(* IEC 61131-3 sources: autonomer-verladearm/plc/codesys, 13 files *)

(* ---- DUT_Pd.st ---- *)
(* Prozessdaten eines MOVITRAC advanced mit MOVIKIT Positioning Drive (Applikationslevel 1, 8 PD).
   Belegung nach Handbuch 33350930 (11/2025), Kap. 8 – im E/A-Abbild des PROFINET-Geräts auf
   diese Felder legen. *)
TYPE ST_PdAxis :
STRUCT
    aPA : ARRAY[1..8] OF WORD;   (* SPS -> Umrichter *)
        (* PA1 Steuerwort, PA2 Geschwindigkeit, PA3 Beschleunigung, PA4 Verzögerung,
           PA5 Ausgänge, PA6 Betriebsart (400 = absolut), PA7/PA8 Zielposition (32 Bit, High/Low) *)
    aPE : ARRAY[1..8] OF WORD;   (* Umrichter -> SPS *)
        (* PE1 Statuswort, PE2 Geschwindigkeit, PE3 Fehlercode, PE4 Moment, PE5 Eingänge,
           PE6 aktive Betriebsart, PE7/PE8 Istposition (32 Bit, High/Low) *)
END_STRUCT
END_TYPE

(* ---- GVL_Achsen.st ---- *)
(* Achsen J1..J3: Prozessdaten (im E/A-Abbild der drei MOVITRAC zuordnen), Fahrbefehle und
   Istwerte. Fahrbefehle schreibt immer nur ein Besitzer (Automatik oder Hand). *)
{attribute 'qualified_only'}
VAR_GLOBAL
    aPd        : ARRAY[1..3] OF ST_PdAxis;   (* E/A-Abbild MOVITRAC J1, J2, J3 *)
    (* Befehle *)
    aCmdZiel   : ARRAY[1..3] OF REAL;        (* ° *)
    aCmdV      : ARRAY[1..3] OF REAL;        (* °/s *)
    aCmdA      : ARRAY[1..3] OF REAL;        (* °/s² *)
    xCmdStart  : BOOL;                       (* Flanke = neues Ziel, halten während der Fahrt *)
    xCmdStop   : BOOL;
    xCmdReset  : BOOL;
    iBesitzer  : INT;                        (* 0 frei, 1 Automatik, 2 Hand *)
    (* Istwerte *)
    aIst       : ARRAY[1..3] OF REAL;        (* ° *)
    xAlleBereit: BOOL;
    xAlleInPos : BOOL;
    xAchsFehler: BOOL;
END_VAR

(* ---- GVL_IO.st ---- *)
(* Ein- und Ausgänge. Im Gerätebaum (TwinCAT: E/A-Abbild der EtherCAT-Klemmen bzw. PROFINET-
   Geräte) diesen Variablen zuordnen. Sicherheitssignale kommen als MELDUNG der Sicherheits-
   steuerung (TwinSAFE) – sie schaltet STO selbst, die SPS kann sie nicht überstimmen.
   Not-Halt am Arm schaltet die Pumpe festverdrahtet über die Sicherheitssteuerung ab (nicht hier). *)
{attribute 'qualified_only'}
VAR_GLOBAL
    (* Bedienung am Schaltschrank *)
    xStartTaster      : BOOL;   (* Leuchttaster "Beladen starten" *)
    xQuittTaster      : BOOL;   (* Quittieren *)
    xBetriebsartHand  : BOOL;   (* Schlüsselschalter: TRUE = Hand, FALSE = Automatik *)
    xLampeStart       : BOOL;   (* Lampe im Starttaster *)
    xMeldeGruen       : BOOL;   (* Park / bereit, Fahrzeug darf fahren *)
    xMeldeGelb        : BOOL;   (* Automatik läuft *)
    xMeldeRot         : BOOL;   (* Störung *)

    (* Handbediengerät (Zustimmung wertet die Sicherheitssteuerung aus) *)
    xHandAchse1       : BOOL;
    xHandAchse2       : BOOL;
    xHandAchse3       : BOOL;
    xHandPlus         : BOOL;
    xHandMinus        : BOOL;
    xHandBremseLueften: BOOL;   (* nur J1/J2, Freigabe zusätzlich durch Sicherheitssteuerung *)

    (* Meldungen der Sicherheitssteuerung *)
    xSicherheitOk     : BOOL;   (* kein Not-Halt, STO aufgehoben *)
    xZustimmung       : BOOL;   (* Zustimmtaster Mittelstellung (nur Hand) *)
    xKlapptreppeRuhe  : BOOL;   (* Klapptreppe in Ruhelage *)
    xLichtschranke    : BOOL;   (* Stellplatz belegt *)

    (* Prozess am Arm *)
    xGrenzNass        : BOOL;   (* Grenzschalter Nachziehen, ca. 10–15 cm über Auslassende: nass *)
    xUeberfuellAus    : BOOL;   (* Überfüllsicherung ausgelöst (schaltet die Pumpe selbst ab) *)
    xKlappeAuf        : BOOL;   (* Absperrklappe Rückmeldung auf *)
    xKlappeZu         : BOOL;   (* Absperrklappe Rückmeldung zu *)
    xKlappeOeffnen    : BOOL;   (* Ausgang Absperrklappe (gehört zum Arm) *)

    (* Abtropfsicherung: rein mechanisch, keine Signale (Entscheidung 04.11.2026) *)

    (* Leitstelle (PLS) – Menge, Pumpe und Füllende steuert die Leitstelle; Signale mit BASF
       abstimmen (Mail an BASF 09.11.2026) *)
    xPlsFreigabe      : BOOL;   (* Verladung freigegeben (Auftrag liegt vor) *)
    iPlsProdukt       : INT;
    aPlsDome          : ARRAY[1..4] OF INT;    (* Füllschritte: DomeNo, 0 = automatisch *)
    iPlsSchritte      : INT;    (* Anzahl Füllschritte (Kammern), 1 = Kammern verbunden *)
    xPlsPumpeLaeuft   : BOOL;   (* Rückmeldung: Pumpe läuft *)
    xPlsBefuellEnde   : BOOL;   (* "Befüllung Ende" für den aktuellen Füllschritt (Pumpe aus) *)
    xArmBereit        : BOOL;   (* an PLS: Arm im Tank, Klappe offen – Befüllung freigegeben *)
    xBefuellStoppen   : BOOL;   (* an PLS: Pumpe abschalten (Störung, Maximalhöhe, Arm am Ende) *)
END_VAR

(* ---- GVL_Param.st ---- *)
(* Parameter Prototyp HETA. Werte aus vision/config/anlagen/heta_prototyp.yaml (drives, arm.joints)
   und docs/fuellstand_ueberfuellsicherung.md. Bei der Inbetriebnahme prüfen. *)
{attribute 'qualified_only'}
VAR_GLOBAL CONSTANT
    INTERFACE_VERSION : INT := 3;
    MAX_WP            : INT := 16;
    TIMEOUT_JOB       : TIME := T#5S;       (* Done muss innerhalb 5 s kommen *)
    TIMEOUT_HEARTBEAT : TIME := T#1S;
    TIMEOUT_MOVE_ADD  : TIME := T#10S;      (* Reserve zur berechneten Fahrzeit *)
    BERUHIGEN         : TIME := T#3S;       (* Auslass pendelt frei aus (J4) *)
    ABTROPFEN         : TIME := T#60S;      (* BASF: 1 min reicht oft nicht – mit Abtropfsicherung *)
    FAKTOR_LANGSAM    : REAL := 0.3;        (* Eintauchen, Herausfahren, Nachziehen *)
    FAKTOR_HAND       : REAL := 0.2;        (* Tippen *)
    TOL_POS           : REAL := 0.2;        (* ° Position erreicht *)
    TOL_PARK          : REAL := 0.5;        (* ° in Parkstellung *)
    MAX_KORREKTUR     : REAL := 50.0;       (* mm Job 2, darüber Abbruch *)
    ANFAHRHOEHE       : REAL := 0.3;        (* m über Domrand (arm.approach_height) *)
    (* Nachziehen mit einem Grenzschalter (Stand 09.11.2026) *)
    SENSOR_HOEHE      : REAL := 0.12;       (* m Grenzschalter über Auslassende (10–15 cm) *)
    NACHZIEH_SCHRITT  : REAL := 0.05;       (* m Hub je Schaltvorgang -> Auslass 7–12 cm unter Spiegel *)
    TROCKEN_ZEIT      : TIME := T#10S;      (* nach dem Hub muss der Grenzschalter trocken sein *)
    MAX_OHNE_SCHALTEN : TIME := T#30M;      (* Pumpe läuft, Grenzschalter schaltet nie: Störung *)
    PUMPE_AUSLAUF     : TIME := T#3S;       (* nach "Pumpe aus" warten, dann Klappe zu *)
    PUMPE_AUS_MAX     : TIME := T#15S;      (* Pumpe meldet nicht aus: Klappe trotzdem zu, Störung *)
END_VAR
VAR_GLOBAL
    (* je Achse J1..J3: Höchstgeschwindigkeit [°/s], Beschleunigung [°/s²], Grenzen und Park [°] *)
    aVmax   : ARRAY[1..3] OF REAL := [6.0, 6.0, 5.93];
    aAmax   : ARRAY[1..3] OF REAL := [1.5, 3.0, 3.95];   (* = vmax / Rampe 4 / 2 / 1,5 s *)
    rRuckzeit : REAL := 0.3;                             (* s, auf allen Achsen gleich *)
    aMin    : ARRAY[1..3] OF REAL := [-120.0, -140.0, -45.0];
    aMax    : ARRAY[1..3] OF REAL := [120.0, 140.0, 45.0];
    aPark   : ARRAY[1..3] OF REAL := [70.0, -135.0, 10.0]; (* heta_prototyp.yaml, bei IBN anpassen *)
    (* Eintauchtiefe je Produkt [m unter Domrand], Index = ProductId 0..9 *)
    (* ca. 20 cm über dem Tankboden: Domrand bis Boden 2,10–2,30 m (BASF 24.11.) – flachster Tank 2,10 m *)
    aEintauchtiefe : ARRAY[0..9] OF REAL := [1.9, 1.9, 1.9, 1.9, 1.9, 1.9, 1.9, 1.9, 1.9, 1.9];
    rMaxHoeheUnterRand : REAL := 0.28;   (* m: Füllende Ebene 2, knapp unter der Überfüllsicherung (ca. 0,2 m) *)
END_VAR

(* ---- GVL_Vision.st ---- *)
(* Schnittstelle Vision-PC <-> SPS, InterfaceVersion 3 (docs/schnittstelle.md).
   Gleiche Namen und Datentypen wie DB_Vision (plc/DB_Vision.db), damit der Vision-Dienst ohne
   Codeänderung verbindet. In der Symbolkonfiguration für OPC UA freigeben (Lesen/Schreiben). *)
{attribute 'qualified_only'}
VAR_GLOBAL
    (* SPS -> PC *)
    HeartbeatPLC   : INT;
    Trigger        : BOOL;
    Job            : INT;      (* 1 messen+planen, 2 nachmessen, 3 Rückfahrt, 0 nur messen *)
    ProductId      : INT;
    DomeNo         : INT;      (* 0 automatisch, n = n-ter offener Dom von vorn *)
    Reset          : BOOL;
    ActualJ1       : REAL;     (* Servo-Istwinkel [°] *)
    ActualJ2       : REAL;
    ActualJ3       : REAL;
    AxesHomed      : BOOL;
    ArmState       : INT;      (* 0 Park, 1 fährt, 2 über Dom, 3 eingetaucht, 9 Störung *)
    (* PC -> SPS *)
    HeartbeatPC    : INT;
    Ready          : BOOL;
    Busy           : BOOL;
    Done           : BOOL;
    Error          : BOOL;
    ErrorCode      : INT;
    ResultId       : DINT;
    TargetX        : REAL;     (* mm, Armbasis *)
    TargetY        : REAL;
    TargetZ        : REAL;
    NormalX        : REAL;
    NormalY        : REAL;
    NormalZ        : REAL;
    DiameterMm     : REAL;
    Confidence     : REAL;
    DomeCount      : INT;
    DomeSelected   : INT;
    WaypointCount  : INT;
    WaypointsJ1    : ARRAY[1..16] OF REAL;   (* Servo-Sollwinkel [°] *)
    WaypointsJ2    : ARRAY[1..16] OF REAL;
    WaypointsJ3    : ARRAY[1..16] OF REAL;
    ApproachIndex  : INT;      (* Stützpunkt "über dem Dom", 0 = keiner *)
    CorrectionX    : REAL;     (* mm, Job 2 *)
    CorrectionY    : REAL;
    InterfaceVersion : INT;
END_VAR

(* ---- F_Hilfen.st ---- *)
(* Hilfsfunktionen für den Ablauf. In CODESYS je Funktion ein eigenes Objekt (POU) anlegen. *)

(* ---------------------------------------------------------------------------------------- *)
(* Arm in Parkstellung? *)
FUNCTION F_InPark : BOOL
VAR
    i : INT;
END_VAR
F_InPark := TRUE;
FOR i := 1 TO 3 DO
    IF ABS(GVL_Achsen.aIst[i] - GVL_Param.aPark[i]) > GVL_Param.TOL_PARK THEN
        F_InPark := FALSE;
    END_IF
END_FOR
END_FUNCTION

(* ---------------------------------------------------------------------------------------- *)
(* Höhe des Auslassendes relativ zum Domrand [m] für eine Lage in der Nachzieh-Tabelle.
   Tabelle = Eintauch-Stützpunkte aus Job 2, gleichmäßig von ANFAHRHOEHE über dem Rand (Lage 1)
   bis rTiefe unter dem Rand (Lage iTab). *)
FUNCTION F_Hoehe : REAL
VAR_INPUT
    rPos   : REAL;   (* 1 .. iTab *)
    iTab   : INT;
    rTiefe : REAL;
END_VAR
IF iTab < 2 THEN
    F_Hoehe := GVL_Param.ANFAHRHOEHE;
ELSE
    F_Hoehe := GVL_Param.ANFAHRHOEHE
               - (rPos - 1.0) / INT_TO_REAL(iTab - 1) * (GVL_Param.ANFAHRHOEHE + rTiefe);
END_IF
END_FUNCTION

(* ---------------------------------------------------------------------------------------- *)
(* Umkehrung: Lage in der Tabelle für eine Höhe relativ zum Domrand. *)
FUNCTION F_PosFuerHoehe : REAL
VAR_INPUT
    rHoehe : REAL;
    iTab   : INT;
    rTiefe : REAL;
END_VAR
IF iTab < 2 THEN
    F_PosFuerHoehe := 1.0;
ELSE
    F_PosFuerHoehe := LIMIT(1.0,
        1.0 + (GVL_Param.ANFAHRHOEHE - rHoehe) / (GVL_Param.ANFAHRHOEHE + rTiefe) * INT_TO_REAL(iTab - 1),
        INT_TO_REAL(iTab));
END_IF
END_FUNCTION

(* ---------------------------------------------------------------------------------------- *)
(* Servowinkel einer Achse für eine Lage in der Tabelle: zwischen den Stützpunkten linear im
   Gelenkraum (wie tools/plc_simulator.py table_at). *)
FUNCTION F_TabWinkel : REAL
VAR_INPUT
    rPos   : REAL;
    iTab   : INT;
    iAchse : INT;
END_VAR
VAR_IN_OUT
    aTab   : ARRAY[1..16, 1..3] OF REAL;
END_VAR
VAR
    k : INT;
    u : REAL;
END_VAR
k := LIMIT(1, DINT_TO_INT(TRUNC(rPos)), MAX(iTab - 1, 1));
u := LIMIT(0.0, rPos - INT_TO_REAL(k), 1.0);
IF iTab < 2 THEN
    F_TabWinkel := aTab[1, iAchse];
ELSE
    F_TabWinkel := aTab[k, iAchse] + u * (aTab[k + 1, iAchse] - aTab[k, iAchse]);
END_IF
END_FUNCTION

(* ---- FB_PdAxis.st ---- *)
(* Eine Achse über MOVIKIT Positioning Drive: Ziel, Geschwindigkeit, Beschleunigung vorgeben,
   Istposition und Status lesen. Positionieren, Rampen und Ruckbegrenzung macht der Umrichter.

   !!! Bitbelegung von Steuer- und Statuswort und die Anwendereinheiten vor der Inbetriebnahme
   mit dem SEW-Handbuch (Kap. 8) und MOVISUITE abgleichen – hier als Konstanten mit
   Platzhalterwerten. Anwendereinheit: 1 Inkrement = 0,001° am Gelenk (in MOVISUITE einstellen). *)
FUNCTION_BLOCK FB_PdAxis
VAR_INPUT
    xEnable  : BOOL;          (* Freigabe (STO aufgehoben, keine Störung) *)
    xStart   : BOOL;          (* steigende Flanke: neues Ziel übernehmen *)
    xStop    : BOOL;          (* Halt mit Verzögerung *)
    xReset   : BOOL;          (* Fehler quittieren *)
    rZiel    : REAL;          (* ° *)
    rV       : REAL;          (* °/s *)
    rA       : REAL;          (* °/s² (Beschleunigung = Verzögerung) *)
END_VAR
VAR_OUTPUT
    rIst     : REAL;          (* ° *)
    xBereit  : BOOL;          (* Umrichter bereit / freigegeben *)
    xInPos   : BOOL;          (* Position erreicht *)
    xFehler  : BOOL;
    wFehler  : WORD;
END_VAR
VAR_IN_OUT
    stPd     : ST_PdAxis;
END_VAR
VAR CONSTANT
    EINHEIT_POS    : REAL := 1000.0;     (* Inkremente je ° (Anwendereinheit 0,001°) *)
    EINHEIT_V      : REAL := 100.0;      (* PA2: 0,01 °/s – prüfen *)
    EINHEIT_A      : REAL := 100.0;      (* PA3/PA4: 0,01 °/s² – prüfen *)
    BETRIEBSART_ABS: WORD := 400;
    (* Steuerwort PA1 – PLATZHALTER, laut Handbuch prüfen *)
    CW_FREIGABE    : WORD := 16#0001;
    CW_START       : WORD := 16#0002;
    CW_HALT        : WORD := 16#0004;
    CW_RESET       : WORD := 16#0100;
    (* Statuswort PE1 – PLATZHALTER, laut Handbuch prüfen *)
    SW_BEREIT      : WORD := 16#0001;
    SW_INPOS       : WORD := 16#0004;
    SW_FEHLER      : WORD := 16#0020;
END_VAR
VAR
    rtStart  : R_TRIG;
    dIst     : DINT;
    dZiel    : DINT;
    wStw     : WORD;
END_VAR

rtStart(CLK := xStart);

(* Istwerte *)
dIst := INT_TO_DINT(WORD_TO_INT(stPd.aPE[7])) * 65536 + WORD_TO_DINT(stPd.aPE[8]);   (* High-Wort mit Vorzeichen *)
rIst := DINT_TO_REAL(dIst) / EINHEIT_POS;
xBereit := (stPd.aPE[1] AND SW_BEREIT) <> 0;
xFehler := (stPd.aPE[1] AND SW_FEHLER) <> 0;
wFehler := stPd.aPE[3];

(* Sollwerte: bei neuem Ziel übernehmen *)
IF rtStart.Q THEN
    dZiel := REAL_TO_DINT(rZiel * EINHEIT_POS);
    stPd.aPA[2] := DINT_TO_WORD(LIMIT(1, REAL_TO_DINT(ABS(rV) * EINHEIT_V), 32767));
    stPd.aPA[3] := DINT_TO_WORD(LIMIT(1, REAL_TO_DINT(ABS(rA) * EINHEIT_A), 32767));
    stPd.aPA[4] := stPd.aPA[3];
    stPd.aPA[7] := DWORD_TO_WORD(SHR(DINT_TO_DWORD(dZiel), 16));
    stPd.aPA[8] := DWORD_TO_WORD(DINT_TO_DWORD(dZiel));
END_IF
stPd.aPA[6] := BETRIEBSART_ABS;

wStw := 0;
IF xEnable THEN wStw := wStw OR CW_FREIGABE; END_IF
IF xEnable AND xStart AND NOT xStop THEN wStw := wStw OR CW_START; END_IF
IF xStop THEN wStw := wStw OR CW_HALT; END_IF
IF xReset THEN wStw := wStw OR CW_RESET; END_IF
stPd.aPA[1] := wStw;

xInPos := ((stPd.aPE[1] AND SW_INPOS) <> 0) AND ABS(rIst - rZiel) <= GVL_Param.TOL_POS;

(* ---- FB_SyncMove.st ---- *)
(* Synchrone Fahrt aller drei Achsen zu einem Stützpunkt (docs/schnittstelle.md):
   Die langsamste Achse bestimmt die Fahrzeit; jede Achse bekommt Geschwindigkeit und
   Beschleunigung proportional zu ihrem Weg, gleiche Ruckzeit auf allen Achsen -> alle starten
   und kommen gleichzeitig an, der Arm fährt die geprüfte Gerade im Gelenkraum.
   Gleiche Rechnung wie Drives.sync() in vision/src/verladearm_vision/drives.py. *)
FUNCTION_BLOCK FB_SyncMove
VAR_INPUT
    xExecute : BOOL;                   (* steigende Flanke startet *)
    aZiel    : ARRAY[1..3] OF REAL;    (* ° *)
    rFaktor  : REAL := 1.0;            (* Geschwindigkeitsfaktor, z. B. 0,3 beim Eintauchen *)
    xAbbruch : BOOL;                   (* Halt mit Verzögerung *)
END_VAR
VAR_OUTPUT
    xBusy    : BOOL;
    xDone    : BOOL;
    xError   : BOOL;
    sFehler  : STRING(80);
    rDauer   : REAL;                   (* s, berechnete Fahrzeit *)
END_VAR
VAR
    rtExec   : R_TRIG;
    iSchritt : INT;
    tonZeit  : TON;
    i        : INT;
    d        : ARRAY[1..3] OF REAL;
    rCruise, rPush, rRamp : REAL;
    rFak     : REAL;
END_VAR

rtExec(CLK := xExecute);
IF rtExec.Q THEN
    xDone := FALSE; xError := FALSE; sFehler := '';
    rFak := LIMIT(0.01, rFaktor, 1.0);
    rCruise := 0.0; rPush := 0.0;
    FOR i := 1 TO 3 DO
        aZiel[i] := LIMIT(GVL_Param.aMin[i], aZiel[i], GVL_Param.aMax[i]);   (* Software-Endlagen *)
        d[i] := ABS(aZiel[i] - GVL_Achsen.aIst[i]);
        rCruise := MAX(rCruise, d[i] / (GVL_Param.aVmax[i] * rFak));
        rPush := MAX(rPush, d[i] / GVL_Param.aAmax[i]);
    END_FOR
    IF rPush < 1.0E-6 THEN
        xDone := TRUE; iSchritt := 0;       (* schon am Ziel *)
    ELSE
        IF SQRT(rPush) >= rCruise THEN      (* Dreieck: Höchstgeschwindigkeit nicht erreicht *)
            rCruise := SQRT(rPush); rRamp := rCruise;
        ELSE
            rRamp := rPush / rCruise;
        END_IF
        rDauer := rCruise + rRamp + GVL_Param.rRuckzeit;
        FOR i := 1 TO 3 DO
            GVL_Achsen.aCmdZiel[i] := aZiel[i];
            GVL_Achsen.aCmdV[i] := MAX(d[i] / rCruise, 0.001);
            GVL_Achsen.aCmdA[i] := MAX(d[i] / rCruise / rRamp, 0.001);
        END_FOR
        GVL_Achsen.xCmdStart := FALSE;      (* ein Zyklus FALSE, damit die Flanke kommt *)
        GVL_Achsen.xCmdStop := FALSE;
        iSchritt := 1;
    END_IF
END_IF

CASE iSchritt OF
1:  GVL_Achsen.xCmdStart := TRUE;
    iSchritt := 2;
2:  (* warten bis alle Achsen am Ziel; Zeitüberwachung *)
    IF xAbbruch THEN
        GVL_Achsen.xCmdStop := TRUE;
        xError := TRUE; sFehler := 'Fahrt abgebrochen'; iSchritt := 0;
    ELSIF GVL_Achsen.xAchsFehler THEN
        xError := TRUE; sFehler := 'Achsfehler (Umrichter)'; iSchritt := 0;
    ELSIF tonZeit.Q THEN
        GVL_Achsen.xCmdStop := TRUE;
        xError := TRUE; sFehler := 'Zeitüberschreitung Fahrt'; iSchritt := 0;
    ELSIF GVL_Achsen.xAlleInPos AND tonZeit.ET > T#200MS THEN
        xDone := TRUE; iSchritt := 0;
    END_IF
END_CASE

tonZeit(IN := iSchritt = 2,
        PT := REAL_TO_TIME(rDauer * 1000.0) + GVL_Param.TIMEOUT_MOVE_ADD);
xBusy := iSchritt <> 0;

(* ---- FB_VisionJob.st ---- *)
(* Auftrag an den Vision-PC (Handshake docs/schnittstelle.md) mit Plausibilitätsprüfung der
   Stützpunkte. Ergebnis bleibt bis zum nächsten Auftrag in den Ausgängen. *)
FUNCTION_BLOCK FB_VisionJob
VAR_INPUT
    xExecute  : BOOL;
    iJob      : INT;
    iProdukt  : INT;
    iDom      : INT;
END_VAR
VAR_OUTPUT
    xBusy     : BOOL;
    xDone     : BOOL;
    xError    : BOOL;
    iFehler   : INT;              (* Fehlercode Vision bzw. 100 + Prüfung SPS *)
    sFehler   : STRING(80);
    iAnzahl   : INT;              (* gültige Stützpunkte *)
    aWp       : ARRAY[1..16, 1..3] OF REAL;
    iUeberDom : INT;              (* ApproachIndex *)
    rDomZ     : REAL;             (* Oberkante Domöffnung [m, Armbasis] *)
    rKorrX, rKorrY : REAL;        (* mm *)
    iDomeCount, iDomeSelected : INT;
END_VAR
VAR
    rtExec    : R_TRIG;
    iSchritt  : INT;
    tonTimeout: TON;
    i, k      : INT;
    aWert     : ARRAY[1..3] OF REAL;
END_VAR

rtExec(CLK := xExecute);
IF rtExec.Q AND iSchritt = 0 THEN
    xDone := FALSE; xError := FALSE; iFehler := 0; sFehler := '';
    iSchritt := 1;
END_IF

CASE iSchritt OF
1:  IF NOT GVL_Vision.Ready THEN
        xError := TRUE; iFehler := 101; sFehler := 'Vision-PC nicht bereit'; iSchritt := 0;
    ELSIF GVL_Vision.InterfaceVersion <> GVL_Param.INTERFACE_VERSION THEN
        xError := TRUE; iFehler := 102; sFehler := 'falsche InterfaceVersion'; iSchritt := 0;
    ELSE
        GVL_Vision.Job := iJob;
        GVL_Vision.ProductId := iProdukt;
        GVL_Vision.DomeNo := iDom;
        GVL_Vision.Trigger := TRUE;
        iSchritt := 2;
    END_IF

2:  IF GVL_Vision.Done THEN
        (* Ergebnis übernehmen *)
        iFehler := GVL_Vision.ErrorCode;
        iAnzahl := LIMIT(0, GVL_Vision.WaypointCount, GVL_Param.MAX_WP);
        FOR i := 1 TO GVL_Param.MAX_WP DO
            aWp[i, 1] := GVL_Vision.WaypointsJ1[i];
            aWp[i, 2] := GVL_Vision.WaypointsJ2[i];
            aWp[i, 3] := GVL_Vision.WaypointsJ3[i];
        END_FOR
        iUeberDom := GVL_Vision.ApproachIndex;
        rDomZ := GVL_Vision.TargetZ / 1000.0;
        rKorrX := GVL_Vision.CorrectionX;
        rKorrY := GVL_Vision.CorrectionY;
        iDomeCount := GVL_Vision.DomeCount;
        iDomeSelected := GVL_Vision.DomeSelected;
        IF GVL_Vision.Error THEN
            xError := TRUE; sFehler := 'Vision-Fehler (Code siehe iFehler)';
        ELSE
            (* Plausibilität: Achsgrenzen jedes Stützpunkts *)
            FOR i := 1 TO iAnzahl DO
                FOR k := 1 TO 3 DO
                    IF aWp[i, k] < GVL_Param.aMin[k] OR aWp[i, k] > GVL_Param.aMax[k] THEN
                        xError := TRUE; iFehler := 103; sFehler := 'Stützpunkt außerhalb der Achsgrenzen';
                    END_IF
                END_FOR
            END_FOR
            IF iJob <> 0 AND iAnzahl = 0 THEN
                xError := TRUE; iFehler := 104; sFehler := 'keine Stützpunkte';
            END_IF
            IF iJob = 2 AND (ABS(rKorrX) > GVL_Param.MAX_KORREKTUR OR ABS(rKorrY) > GVL_Param.MAX_KORREKTUR) THEN
                xError := TRUE; iFehler := 105; sFehler := 'Korrektur Job 2 zu groß';
            END_IF
        END_IF
        GVL_Vision.Trigger := FALSE;
        iSchritt := 3;
    ELSIF tonTimeout.Q THEN
        GVL_Vision.Trigger := FALSE;
        xError := TRUE; iFehler := 106; sFehler := 'Zeitüberschreitung Vision-PC';
        iSchritt := 0;
    END_IF

3:  IF NOT GVL_Vision.Done THEN      (* PC hat Done gelöscht *)
        xDone := NOT xError;
        iSchritt := 0;
    ELSIF tonTimeout.Q THEN
        xError := TRUE; iFehler := 107; sFehler := 'Done wird nicht gelöscht'; iSchritt := 0;
    END_IF
END_CASE

tonTimeout(IN := iSchritt = 2 OR iSchritt = 3, PT := GVL_Param.TIMEOUT_JOB);
xBusy := iSchritt <> 0;

(* ---- PRG_Achsen.st ---- *)
(* Jeden Zyklus: drei Achsen bedienen, Istwerte an den Vision-PC. Vor PRG_Main aufrufen. *)
PROGRAM PRG_Achsen
VAR
    fbAchse : ARRAY[1..3] OF FB_PdAxis;
    i       : INT;
END_VAR

GVL_Achsen.xAlleBereit := TRUE;
GVL_Achsen.xAlleInPos := TRUE;
GVL_Achsen.xAchsFehler := FALSE;
FOR i := 1 TO 3 DO
    fbAchse[i](
        xEnable := GVL_IO.xSicherheitOk,
        xStart  := GVL_Achsen.xCmdStart,
        xStop   := GVL_Achsen.xCmdStop,
        xReset  := GVL_Achsen.xCmdReset,
        rZiel   := GVL_Achsen.aCmdZiel[i],
        rV      := GVL_Achsen.aCmdV[i],
        rA      := GVL_Achsen.aCmdA[i],
        stPd    := GVL_Achsen.aPd[i]);
    GVL_Achsen.aIst[i] := fbAchse[i].rIst;
    GVL_Achsen.xAlleBereit := GVL_Achsen.xAlleBereit AND fbAchse[i].xBereit;
    GVL_Achsen.xAlleInPos := GVL_Achsen.xAlleInPos AND fbAchse[i].xInPos;
    GVL_Achsen.xAchsFehler := GVL_Achsen.xAchsFehler OR fbAchse[i].xFehler;
END_FOR

(* Multiturn-Absolutgeber: Lage gilt sofort, keine Referenzfahrt *)
GVL_Vision.ActualJ1 := GVL_Achsen.aIst[1];
GVL_Vision.ActualJ2 := GVL_Achsen.aIst[2];
GVL_Vision.ActualJ3 := GVL_Achsen.aIst[3];
GVL_Vision.AxesHomed := GVL_Achsen.xAlleBereit AND NOT GVL_Achsen.xAchsFehler;

(* ---- PRG_Hand.st ---- *)
(* Handbetrieb (Schlüsselschalter Hand) mit dem Handbediengerät: eine Achse wählen, mit + / −
   tippen, solange Zustimmtaster (Mittelstellung) gehalten wird. Reduzierte Geschwindigkeit,
   Software-Endlagen bleiben aktiv. Zustimmung und Not-Halt wertet die Sicherheitssteuerung aus;
   hier nur die Bewegung.

   Bremse lüften (nur J1/J2, Arm von Hand schieben): Antrieb in STO, Bremse über den
   Bremsausgang des Umrichters öffnen – Funktion und Freigabe bei SEW/Sicherheitskonzept klären.
   J3 nie lüften (Selbsthemmung nicht zugesichert). *)
PROGRAM PRG_Hand
VAR
    iAchse   : INT;
    xFahrt   : BOOL;
    i        : INT;
END_VAR

IF NOT GVL_IO.xBetriebsartHand OR PRG_Main.iSchritt <> 0 AND PRG_Main.iSchritt < 900 THEN
    xFahrt := FALSE;
    RETURN;
END_IF

iAchse := 0;
IF GVL_IO.xHandAchse1 THEN iAchse := 1;
ELSIF GVL_IO.xHandAchse2 THEN iAchse := 2;
ELSIF GVL_IO.xHandAchse3 THEN iAchse := 3;
END_IF

IF iAchse > 0 AND GVL_IO.xZustimmung AND GVL_IO.xSicherheitOk
   AND (GVL_IO.xHandPlus XOR GVL_IO.xHandMinus) THEN
    IF NOT xFahrt THEN
        (* Ziel = Endlage in Tipprichtung, andere Achsen bleiben stehen *)
        FOR i := 1 TO 3 DO
            GVL_Achsen.aCmdZiel[i] := GVL_Achsen.aIst[i];
            GVL_Achsen.aCmdV[i] := 0.001;
            GVL_Achsen.aCmdA[i] := 0.001;
        END_FOR
        GVL_Achsen.aCmdZiel[iAchse] := SEL(GVL_IO.xHandPlus, GVL_Param.aMin[iAchse], GVL_Param.aMax[iAchse]);
        GVL_Achsen.aCmdV[iAchse] := GVL_Param.aVmax[iAchse] * GVL_Param.FAKTOR_HAND;
        GVL_Achsen.aCmdA[iAchse] := GVL_Param.aAmax[iAchse];
        GVL_Achsen.iBesitzer := 2;
        GVL_Achsen.xCmdStop := FALSE;
        GVL_Achsen.xCmdStart := FALSE;   (* Flanke im nächsten Zyklus *)
        xFahrt := TRUE;
    ELSE
        GVL_Achsen.xCmdStart := TRUE;
    END_IF
ELSIF xFahrt THEN
    (* losgelassen: anhalten *)
    GVL_Achsen.xCmdStart := FALSE;
    GVL_Achsen.xCmdStop := TRUE;
    xFahrt := FALSE;
ELSE
    GVL_Achsen.xCmdStop := TRUE;      (* steht: Halt bleibt aktiv, Automatik nimmt ihn beim Start zurück *)
    GVL_Achsen.iBesitzer := 0;
END_IF

(* ---- PRG_Heartbeat.st ---- *)
(* Heartbeat SPS -> PC alle 100 ms, Überwachung des PC-Heartbeats (Ausfall > 1 s). *)
PROGRAM PRG_Heartbeat
VAR
    tonTakt   : TON;
    tonPc     : TON;
    iLetzter  : INT;
END_VAR
VAR_OUTPUT
    xPcOk     : BOOL;     (* PC-Heartbeat läuft *)
END_VAR

tonTakt(IN := NOT tonTakt.Q, PT := T#100MS);
IF tonTakt.Q THEN
    IF GVL_Vision.HeartbeatPLC >= 32766 THEN
        GVL_Vision.HeartbeatPLC := 0;
    ELSE
        GVL_Vision.HeartbeatPLC := GVL_Vision.HeartbeatPLC + 1;
    END_IF
END_IF

tonPc(IN := GVL_Vision.HeartbeatPC = iLetzter, PT := GVL_Param.TIMEOUT_HEARTBEAT);
iLetzter := GVL_Vision.HeartbeatPC;
xPcOk := NOT tonPc.Q;

(* ---- PRG_Main.st ---- *)
(* Automatischer Verladeablauf – entspricht tools/plc_simulator.py (sequence, fill_tank).
   Je Füllschritt (Kammer): Job 1 -> über den Dom -> Job 2 -> eintauchen -> Klappe auf, "Arm
   bereit" -> Befüllung durch die Leitstelle, Nachziehen über einen Grenzschalter -> Pumpe aus,
   Klappe zu, abtropfen -> heraus -> nächste Kammer (Job 1 vom Dom aus) oder Job 3 -> Park.
   Die Abtropfsicherung arbeitet rein mechanisch (keine Signale).

   Menge, Pumpe und Füllende steuert die Leitstelle. Schutzebenen
   (docs/fuellstand_ueberfuellsicherung.md):
   1. Leitstelle meldet "Befüllung Ende" (Pumpe aus),
   2. Maximalhöhe aus Armhöhe + Grenzschalter bzw. Arm kann nicht weiter nachziehen
      -> "Befüllung stoppen" an die Leitstelle,
   3. Überfüllsicherung – letzte Ebene, schaltet die Pumpe selbst ab; hier nur Störung.
   Reihenfolge immer: erst Pumpe aus (Rückmeldung + Auslaufzeit), dann Klappe zu.

   Muster: Bausteine werden je Zyklus genau einmal VOR dem CASE aufgerufen. Ein Schritt setzt
   den Startmerker, der nächste Schritt wartet auf Done/Error und nimmt den Merker zurück. *)
PROGRAM PRG_Main
VAR_OUTPUT
    iSchritt    : INT;
    sMeldung    : STRING(80);
END_VAR
VAR
    iKammer     : INT;                 (* Füllschritt 1..iPlsSchritte *)
    iWp         : INT;                 (* aktueller Stützpunkt *)
    fbJob       : FB_VisionJob;
    fbMove      : FB_SyncMove;
    xJobStart   : BOOL;
    iJobNr      : INT;
    iDomNr      : INT;
    xMoveStart  : BOOL;
    aZiel       : ARRAY[1..3] OF REAL;
    rFaktor     : REAL := 1.0;
    xWarten     : BOOL;
    tWarte      : TIME;
    tonWarte    : TON;
    rtStart     : R_TRIG;
    rtQuitt     : R_TRIG;
    (* Nachzieh-Tabelle aus Job 2 *)
    aTab        : ARRAY[1..16, 1..3] OF REAL;
    iTab        : INT;
    rTiefe      : REAL;                (* m unter Domrand *)
    rPosTab     : REAL;                (* 1 = Anfahrpunkt, iTab = eingetaucht *)
    rHoehe      : REAL;                (* Auslassende relativ zum Domrand [m] *)
    rSpiegel    : REAL;                (* Spiegel relativ zum Domrand [m] *)
    xNachStoppStoerung : BOOL;         (* nach dem Pumpenstopp in die Störung statt abtropfen *)
    tonTrocken  : TON;                 (* nach dem Hub muss der Grenzschalter trocken sein *)
    tonOhneSchalten : TON;             (* Pumpe läuft, Grenzschalter schaltet nicht *)
    tonPumpeAus : TON;                 (* Warten auf "Pumpe aus" *)
    tonAuslauf  : TON;                 (* Auslaufzeit der Pumpe *)
    xAuto       : BOOL;
    i           : INT;
END_VAR

rtStart(CLK := GVL_IO.xStartTaster);
rtQuitt(CLK := GVL_IO.xQuittTaster);

(* Bausteine: einmal je Zyklus *)
fbJob(xExecute := xJobStart, iJob := iJobNr, iProdukt := GVL_IO.iPlsProdukt, iDom := iDomNr);
fbMove(xExecute := xMoveStart, aZiel := aZiel, rFaktor := rFaktor, xAbbruch := iSchritt >= 900);
tonWarte(IN := xWarten, PT := tWarte);
tonTrocken(IN := iSchritt = 56, PT := GVL_Param.TROCKEN_ZEIT);
tonOhneSchalten(IN := iSchritt = 51 AND GVL_IO.xPlsPumpeLaeuft AND NOT GVL_IO.xGrenzNass,
                PT := GVL_Param.MAX_OHNE_SCHALTEN);
tonPumpeAus(IN := (iSchritt = 58 OR iSchritt = 900) AND GVL_IO.xPlsPumpeLaeuft,
            PT := GVL_Param.PUMPE_AUS_MAX);
tonAuslauf(IN := (iSchritt = 58 OR iSchritt = 900) AND NOT GVL_IO.xPlsPumpeLaeuft,
           PT := GVL_Param.PUMPE_AUSLAUF);

(* Verriegelungen während der Automatik *)
xAuto := GVL_IO.xSicherheitOk AND GVL_IO.xKlapptreppeRuhe AND PRG_Heartbeat.xPcOk
         AND NOT GVL_IO.xBetriebsartHand;
IF iSchritt > 0 AND iSchritt < 900 THEN
    IF NOT xAuto OR (NOT GVL_IO.xLichtschranke AND iSchritt < 80) THEN   (* bei Rückfahrt darf das Fahrzeug weg sein *)
        sMeldung := 'Verriegelung: Sicherheit, Treppe, Lichtschranke, PC oder Betriebsart';
        iSchritt := 900;
    ELSIF GVL_IO.xUeberfuellAus THEN
        sMeldung := 'Überfüllsicherung ausgelöst';
        iSchritt := 900;
    END_IF
END_IF

CASE iSchritt OF
0:  (* bereit *)
    GVL_Vision.ArmState := 0;
    GVL_Achsen.iBesitzer := 0;
    GVL_IO.xKlappeOeffnen := FALSE; GVL_IO.xArmBereit := FALSE; GVL_IO.xBefuellStoppen := FALSE;
    IF rtStart.Q AND F_InPark() AND xAuto AND GVL_IO.xLichtschranke AND GVL_IO.xPlsFreigabe
       AND GVL_Vision.Ready AND GVL_Vision.AxesHomed AND GVL_IO.iPlsSchritte >= 1 THEN
        GVL_Achsen.iBesitzer := 1;
        iKammer := 1;
        sMeldung := '';
        iSchritt := 10;
    END_IF

(* --- Job 1: Dom messen, Bahn planen ------------------------------------------------------- *)
10: iJobNr := 1; iDomNr := GVL_IO.aPlsDome[iKammer]; xJobStart := TRUE; iSchritt := 11;
11: IF fbJob.xDone THEN
        xJobStart := FALSE; iWp := 1; GVL_Vision.ArmState := 1; iSchritt := 20;
    ELSIF fbJob.xError THEN
        xJobStart := FALSE; sMeldung := CONCAT('Job 1: ', fbJob.sFehler); iSchritt := 900;
    END_IF

(* --- Stützpunkte bis über den Dom --------------------------------------------------------- *)
20: FOR i := 1 TO 3 DO aZiel[i] := fbJob.aWp[iWp, i]; END_FOR
    rFaktor := 1.0; xMoveStart := TRUE; iSchritt := 21;
21: IF fbMove.xDone THEN
        xMoveStart := FALSE;
        IF iWp < fbJob.iUeberDom THEN
            iWp := iWp + 1; iSchritt := 20;
        ELSE
            GVL_Vision.ArmState := 2; tWarte := GVL_Param.BERUHIGEN; xWarten := TRUE; iSchritt := 25;
        END_IF
    ELSIF fbMove.xError THEN
        xMoveStart := FALSE; sMeldung := fbMove.sFehler; iSchritt := 900;
    END_IF
25: IF tonWarte.Q THEN xWarten := FALSE; iSchritt := 30; END_IF

(* --- Job 2: Auslass nachmessen, Eintauch-Stützpunkte = Nachzieh-Tabelle ------------------- *)
30: iJobNr := 2; xJobStart := TRUE; iSchritt := 31;
31: IF fbJob.xDone THEN
        xJobStart := FALSE;
        iTab := fbJob.iAnzahl;
        FOR iWp := 1 TO iTab DO
            FOR i := 1 TO 3 DO aTab[iWp, i] := fbJob.aWp[iWp, i]; END_FOR
        END_FOR
        rTiefe := GVL_Param.aEintauchtiefe[LIMIT(0, GVL_IO.iPlsProdukt, 9)];
        iWp := 1; iSchritt := 40;
    ELSIF fbJob.xError THEN
        xJobStart := FALSE; sMeldung := CONCAT('Job 2: ', fbJob.sFehler); iSchritt := 80;
    END_IF

(* --- Eintauchen: Anfahrpunkt normal, danach langsam --------------------------------------- *)
40: FOR i := 1 TO 3 DO aZiel[i] := aTab[iWp, i]; END_FOR
    rFaktor := SEL(iWp = 1, GVL_Param.FAKTOR_LANGSAM, 1.0);
    xMoveStart := TRUE; iSchritt := 41;
41: IF fbMove.xDone THEN
        xMoveStart := FALSE;
        IF iWp < iTab THEN
            iWp := iWp + 1; iSchritt := 40;
        ELSE
            rPosTab := INT_TO_REAL(iTab);
            GVL_Vision.ArmState := 3;
            xNachStoppStoerung := FALSE;
            iSchritt := 50;
        END_IF
    ELSIF fbMove.xError THEN
        xMoveStart := FALSE; sMeldung := fbMove.sFehler; iSchritt := 900;
    END_IF

(* --- Klappe auf, "Arm bereit" an die Leitstelle -------------------------------------------- *)
50: GVL_IO.xKlappeOeffnen := TRUE; GVL_IO.xBefuellStoppen := FALSE;
    IF GVL_IO.xKlappeAuf THEN GVL_IO.xArmBereit := TRUE; iSchritt := 51; END_IF

(* --- Befüllung durch die Leitstelle, Nachziehen über einen Grenzschalter ------------------ *)
51: rHoehe := F_Hoehe(rPosTab, iTab, rTiefe);
    IF GVL_IO.xPlsBefuellEnde THEN                                  (* Ebene 1: Leitstelle *)
        sMeldung := 'Leitstelle: Befüllung Ende'; iSchritt := 58;
    ELSIF tonOhneSchalten.Q THEN
        sMeldung := 'Grenzschalter schaltet nicht (Pumpe läuft zu lange)';
        xNachStoppStoerung := TRUE; iSchritt := 58;
    ELSIF GVL_IO.xGrenzNass THEN                                    (* Spiegel auf Sensorhöhe *)
        rSpiegel := rHoehe + GVL_Param.SENSOR_HOEHE;
        IF rSpiegel >= -GVL_Param.rMaxHoeheUnterRand THEN
            sMeldung := 'Maximalhöhe erreicht – Befüllung stoppen'; iSchritt := 58;   (* Ebene 2 *)
        ELSIF rPosTab <= 1.0 THEN
            sMeldung := 'Arm kann nicht weiter nachziehen – Befüllung stoppen'; iSchritt := 58;
        ELSE                                                        (* Hub um NACHZIEH_SCHRITT *)
            rPosTab := F_PosFuerHoehe(rHoehe + GVL_Param.NACHZIEH_SCHRITT, iTab, rTiefe);
            FOR i := 1 TO 3 DO aZiel[i] := F_TabWinkel(rPosTab, iTab, i, aTab); END_FOR
            rFaktor := GVL_Param.FAKTOR_LANGSAM; xMoveStart := TRUE;
            iSchritt := 55;
        END_IF
    END_IF
55: (* Nachziehen läuft, Klappe bleibt auf, Pumpe läuft weiter *)
    IF fbMove.xDone THEN
        xMoveStart := FALSE; iSchritt := 56;
    ELSIF fbMove.xError THEN
        xMoveStart := FALSE; sMeldung := fbMove.sFehler; iSchritt := 900;
    END_IF
56: (* nach dem Hub muss der Grenzschalter trocken werden *)
    IF NOT GVL_IO.xGrenzNass THEN
        iSchritt := 51;
    ELSIF tonTrocken.Q THEN
        sMeldung := 'Grenzschalter nach dem Nachziehen weiter nass (Belag/Defekt)';
        xNachStoppStoerung := TRUE; iSchritt := 58;
    ELSIF GVL_IO.xPlsBefuellEnde THEN
        sMeldung := 'Leitstelle: Befüllung Ende'; iSchritt := 58;
    END_IF

(* --- erst Pumpe aus (Leitstelle), dann Klappe zu ----------------------------------------- *)
58: GVL_IO.xArmBereit := FALSE;
    GVL_IO.xBefuellStoppen := TRUE;                                 (* bei "Ende" ohnehin aus *)
    IF tonAuslauf.Q THEN
        iSchritt := 60;
    ELSIF tonPumpeAus.Q THEN
        sMeldung := 'Pumpe meldet nicht aus – Klappe zu'; xNachStoppStoerung := TRUE; iSchritt := 60;
    END_IF

(* --- Klappe zu, abtropfen ----------------------------------------------------------------- *)
60: GVL_IO.xKlappeOeffnen := FALSE; GVL_IO.xArmBereit := FALSE;
    IF GVL_IO.xKlappeZu THEN
        GVL_IO.xBefuellStoppen := FALSE;
        IF xNachStoppStoerung THEN
            iSchritt := 900;
        ELSE
            tWarte := GVL_Param.ABTROPFEN; xWarten := TRUE; iSchritt := 62;
        END_IF
    END_IF
62: IF tonWarte.Q THEN xWarten := FALSE; iSchritt := 65; END_IF

(* --- senkrecht heraus bis zum Anfahrpunkt ------------------------------------------------- *)
65: rPosTab := 1.0;
    FOR i := 1 TO 3 DO aZiel[i] := aTab[1, i]; END_FOR
    rFaktor := GVL_Param.FAKTOR_LANGSAM; xMoveStart := TRUE; iSchritt := 66;
66: IF fbMove.xDone THEN
        xMoveStart := FALSE; GVL_Vision.ArmState := 2; iSchritt := 70;
    ELSIF fbMove.xError THEN
        xMoveStart := FALSE; sMeldung := fbMove.sFehler; iSchritt := 900;
    END_IF

(* --- nächste Kammer oder Rückfahrt ------------------------------------------------------- *)
70: IF iKammer < GVL_IO.iPlsSchritte THEN
        iKammer := iKammer + 1; iSchritt := 10;
    ELSE
        iSchritt := 80;
    END_IF

(* --- Job 3: Rückfahrt in die Parkstellung ------------------------------------------------- *)
80: GVL_IO.xKlappeOeffnen := FALSE; GVL_IO.xArmBereit := FALSE;
    GVL_Achsen.iBesitzer := 1;
    iJobNr := 3; iDomNr := 0; xJobStart := TRUE; iSchritt := 81;
81: IF fbJob.xDone THEN
        xJobStart := FALSE; iWp := 1; GVL_Vision.ArmState := 1; iSchritt := 85;
    ELSIF fbJob.xError THEN
        xJobStart := FALSE; sMeldung := CONCAT('Job 3: ', fbJob.sFehler); iSchritt := 900;
    END_IF
85: FOR i := 1 TO 3 DO aZiel[i] := fbJob.aWp[iWp, i]; END_FOR
    rFaktor := SEL(iWp <= 2, 1.0, GVL_Param.FAKTOR_LANGSAM);     (* erst langsam heraus *)
    xMoveStart := TRUE; iSchritt := 86;
86: IF fbMove.xDone THEN
        xMoveStart := FALSE;
        IF iWp < fbJob.iAnzahl THEN
            iWp := iWp + 1; iSchritt := 85;
        ELSE
            GVL_Vision.ArmState := 0; GVL_Achsen.iBesitzer := 0;
            sMeldung := 'Parkstellung – Fahrzeug darf wegfahren'; iSchritt := 0;
        END_IF
    ELSIF fbMove.xError THEN
        xMoveStart := FALSE; sMeldung := fbMove.sFehler; iSchritt := 900;
    END_IF

(* --- Störung ------------------------------------------------------------------------------ *)
900: GVL_Achsen.xCmdStop := TRUE;
    (* Störung: Pumpe abschalten lassen, Klappe erst nach Pumpe aus (bzw. nach PUMPE_AUS_MAX) zu *)
    GVL_IO.xArmBereit := FALSE;
    GVL_IO.xBefuellStoppen := GVL_IO.xPlsPumpeLaeuft OR NOT GVL_IO.xKlappeZu;
    IF tonAuslauf.Q OR tonPumpeAus.Q OR NOT GVL_IO.xKlappeAuf THEN
        GVL_IO.xKlappeOeffnen := FALSE;
    END_IF
    GVL_Vision.ArmState := 9;
    xJobStart := FALSE; xMoveStart := FALSE; xWarten := FALSE;
    GVL_Achsen.xCmdReset := GVL_IO.xQuittTaster;
    IF rtQuitt.Q THEN iSchritt := 910; END_IF
910: (* quittiert: Start = "Automatisch in Parkstellung" (Job 3) oder Handbetrieb *)
    GVL_Achsen.xCmdStop := FALSE; GVL_Achsen.xCmdReset := FALSE;
    GVL_Achsen.iBesitzer := 0;
    GVL_IO.xKlappeOeffnen := FALSE;
    GVL_IO.xBefuellStoppen := GVL_IO.xPlsPumpeLaeuft;
    IF F_InPark() THEN
        GVL_Vision.ArmState := 0; iSchritt := 0;
    ELSIF rtStart.Q AND GVL_IO.xSicherheitOk AND NOT GVL_IO.xBetriebsartHand THEN
        iSchritt := 80;
    END_IF
END_CASE

(* Leuchtmelder *)
GVL_IO.xMeldeRot := iSchritt >= 900;
GVL_IO.xMeldeGelb := iSchritt > 0 AND iSchritt < 900;
GVL_IO.xMeldeGruen := iSchritt = 0 AND F_InPark();
GVL_IO.xLampeStart := iSchritt = 0 AND F_InPark() AND GVL_IO.xPlsFreigabe;
